(*
SPDX-FileCopyrightText: © 2026 Oleksandr Tiutyk <trofimich@gmail.com>
SPDX-License-Identifier: MIT
License: https://opensource.org/license/mit
*)

(*!
<summary>Provides STRING constants and helpers for text manipulation and value formatting.</summary>
<description>
Buffer ownership and size requirements are defined by each operation. ANY formatting reads the caller's value
through its type descriptor. Try methods contain exceptions; this does not validate buffer lifetime or undo
partial modifications.
Runtime type diagnostics use TYPE_ names for known classes and decimal codes for unknown values.
</description>
*)

{attribute 'no_explicit_call' := 'Direct call is not allowed'}
PROGRAM Strings
VAR_INPUT CONSTANT
	CharSize : BYTE := 1;
	//! <summary>ASCII space byte; values below it are control bytes in lexical text filters.</summary>
	ASCII_SPACE : BYTE := BYTE#16#20;
	NewLine : STRING(1) := '$R';
	Empty : STRING(0) := '';
	//! <summary>Standard three-dot ellipsis sequence for single-byte text truncation.</summary>
	ELLIPSIS : STRING(3) := '...';
END_VAR
VAR
	{attribute 'hide'} 
	_ClassName : STRING := __POUNAME();
END_VAR

(*!
<summary>Formats a supported ANY value as text of at most 255 characters.</summary>
<description>
Reads the borrowed live payload of supported types. Unsupported type classes produce a diagnostic marker
containing the type and size instead of interpreting the payload. The result is an independent bounded value.
</description>
*)
METHOD AnyToString : STRING(255)
VAR_INPUT
	value : ANY;
END_VAR
AnyToString := InternalAnyToString255(value := value);
END_METHOD

(*!
<summary>Formats a supported ANY value as text of at most 255 characters.</summary>
<description>
Reads the borrowed live payload of supported types. Unsupported type classes produce a diagnostic marker
containing the type and size instead of interpreting the payload. The result is an independent bounded value.
</description>
*)
METHOD AnyToString255 : STRING(255)
VAR_INPUT
	value : ANY;
END_VAR
AnyToString255 := InternalAnyToString255(value := value);
END_METHOD

(*!
<summary>
Formats a supported ANY value as text of at most 255 characters, fitting longer strings with an ellipsis
('...').
</summary>
<description>
Reads the borrowed live payload of supported types. String values longer than 255 characters are truncated to
252 characters and end with '...'. Non-string types and strings fitting in 255 characters are formatted
identically to AnyToString255.
</description>
<param name="value">Borrowed live value to format.</param>
*)
METHOD AnyToStringFit255 : STRING(255)
VAR_INPUT
	value : ANY;
END_VAR
VAR
	valueLength : UDINT;
END_VAR
AnyToStringFit255 := InternalAnyToString255(value := value);

IF value.TypeClass = __SYSTEM.TYPE_CLASS.TYPE_STRING THEN
	valueLength := InternalGetLength(value := value.pValue);

	IF valueLength > 255 THEN
		AnyToStringFit255 := Tc2_Standard.CONCAT(STR1 := Tc2_Standard.LEFT(STR := AnyToStringFit255, SIZE := 252), STR2 := '...');
	END_IF
ELSIF value.TypeClass = __SYSTEM.TYPE_CLASS.TYPE_WSTRING THEN
	valueLength := WideStrings.InternalGetLength(value := value.pValue);

	IF valueLength > 255 THEN
		AnyToStringFit255 := Tc2_Standard.CONCAT(STR1 := Tc2_Standard.LEFT(STR := AnyToStringFit255, SIZE := 252), STR2 := '...');
	END_IF
END_IF
END_METHOD

(*!
<summary>Appends one STRING to a caller-owned STRING buffer.</summary>
<description>
Requires live, null-terminated strings and a writable target whose declared size describes its capacity. After
validating the target type, an empty source completes without modifying the target. A non-STRING target raises
NotSupportedException; failure of the append helper raises TargetVariableMemoryOverflowException. Source
storage is borrowed only for this call.
Known runtime type classes appear by their TYPE_ names; unknown values retain their decimal codes.
</description>
*)
//!<param name="targetString">Writable STRING buffer to append to.</param>
//!<param name="sourceString">Text to append; empty leaves the target unchanged.</param>
METHOD Append
VAR_INPUT
	targetString : ANY_STRING;
END_VAR
VAR_IN_OUT CONSTANT
	sourceString : STRING;
END_VAR
VAR
	formattedExceptionMessage : WSTRING(255);
	
END_VAR
IF targetString.TypeClass <> __SYSTEM.TYPE_CLASS.TYPE_STRING THEN
	formattedExceptionMessage := Tc2_Utilities.WCONCAT(
		STR1 := "Not supported type ",
		STR2 := SystemTypeClassConvertor.ToWideString(typeClass := targetString.TypeClass)
	);

	Exceptions.ThrowNotSupported(
		sourceNamespaceName := NamespaceName,
		sourceClassName := ClassName,
		sourcePOUName := __POUNAME(),
		sourcePosition := __POSITION(),
		message := formattedExceptionMessage
	);
END_IF

IF sourceString = '' THEN
	RETURN;
END_IF

IF NOT InternalAppend(
	targetString := targetString,
	sourceString1 := ADR(sourceString),
	sourceString2 := 0,
	sourceString3 := 0,
	sourceString4 := 0,
	sourceString5 := 0,
	sourceString6 := 0,
	sourceString7 := 0,
	sourceString8 := 0,
	sourceString9 := 0,
	sourceString10 := 0
) THEN
	Exceptions.ThrowTargetVariableMemoryOverflow(
		sourceNamespaceName := NamespaceName,
		sourceClassName := ClassName,
		sourcePOUName := __POUNAME(),
		sourcePosition := __POSITION(),
		targetVariableName := 'targetString',
		targetVariableSize := TO_ULINT(targetString.diSize)
	); 
END_IF
END_METHOD

(*!
<summary>Appends up to ten STRING fragments in argument order, skipping empty fragments.</summary>
<description>
Requires live, null-terminated source strings and a writable STRING target with valid capacity metadata. Empty
fragments do not stop processing; if all are empty, the target is unchanged and the operation succeeds. Raises
NotSupportedException for a non-STRING target or TargetVariableMemoryOverflowException when appending fails.
Processing stops on the first append failure; earlier modifications are not rolled back. Source storage is
borrowed only for this call.
Known runtime type classes appear by their TYPE_ names; unknown values retain their decimal codes.
</description>
*)
METHOD Append255
VAR_INPUT
	targetString : ANY_STRING;
	sourceString1 : STRING(255);
	sourceString2 : STRING(255) := '';
	sourceString3 : STRING(255) := '';
	sourceString4 : STRING(255) := '';
	sourceString5 : STRING(255) := '';
	sourceString6 : STRING(255) := '';
	sourceString7 : STRING(255) := '';
	sourceString8 : STRING(255) := '';
	sourceString9 : STRING(255) := '';
	sourceString10 : STRING(255) := '';
END_VAR
VAR
	formattedExceptionMessage : WSTRING(255);
	
END_VAR
IF targetString.TypeClass <> __SYSTEM.TYPE_CLASS.TYPE_STRING THEN
	formattedExceptionMessage := Tc2_Utilities.WCONCAT(
		STR1 := "Not supported type ",
		STR2 := SystemTypeClassConvertor.ToWideString(typeClass := targetString.TypeClass)
	);

	Exceptions.ThrowNotSupported(
		sourceNamespaceName := NamespaceName,
		sourceClassName := ClassName,
		sourcePOUName := __POUNAME(),
		sourcePosition := __POSITION(),
		message := formattedExceptionMessage
	);
END_IF

	IF NOT InternalAppend(
		targetString := targetString,
		sourceString1 := ADR(sourceString1),
		sourceString2 := ADR(sourceString2),
		sourceString3 := ADR(sourceString3),
		sourceString4 := ADR(sourceString4),
		sourceString5 := ADR(sourceString5),
		sourceString6 := ADR(sourceString6),
		sourceString7 := ADR(sourceString7),
		sourceString8 := ADR(sourceString8),
		sourceString9 := ADR(sourceString9),
		sourceString10 := ADR(sourceString10)
	) THEN
	Exceptions.ThrowTargetVariableMemoryOverflow(
		sourceNamespaceName := NamespaceName,
		sourceClassName := ClassName,
		sourcePOUName := __POUNAME(),
		sourcePosition := __POSITION(),
		targetVariableName := 'targetString',
		targetVariableSize := TO_ULINT(targetString.diSize)
	); 
END_IF
END_METHOD

(*!
<summary>
Appends one STRING to a caller-owned STRING buffer, fitting available capacity with an ellipsis ('...') if
exceeded.
</summary>
<description>
Requires a writable STRING target with valid capacity metadata. If the appended text exceeds target capacity,
it is truncated so the final characters are '...' followed by a null-terminator. Raises NotSupportedException
for a non-STRING target. Source storage is borrowed only for this call.
Known runtime type classes appear by their TYPE_ names; unknown values retain their decimal codes.
</description>
<param name="targetString">Writable STRING buffer to append to.</param>
<param name="sourceString">Text to append; empty leaves the target unchanged.</param>
*)
METHOD AppendFit
VAR_INPUT
	targetString : ANY_STRING;
END_VAR
VAR_IN_OUT CONSTANT
	sourceString : STRING;
END_VAR
VAR
	formattedExceptionMessage : WSTRING(255);
END_VAR
IF targetString.TypeClass <> __SYSTEM.TYPE_CLASS.TYPE_STRING THEN
	formattedExceptionMessage := WideStrings.Concat255(
		"Not supported type ",
		SystemTypeClassConvertor.ToWideString(typeClass := targetString.TypeClass)
	);

	Exceptions.ThrowNotSupported(
		sourceNamespaceName := NamespaceName,
		sourceClassName := ClassName,
		sourcePOUName := __POUNAME(),
		sourcePosition := __POSITION(),
		message := formattedExceptionMessage
	);
END_IF

InternalAppendFit(targetString := targetString, sourceString := ADR(sourceString));
END_METHOD

(*!
<summary>
Appends up to ten STRING fragments in argument order, fitting available capacity with an ellipsis ('...') if
exceeded.
</summary>
<description>
Requires a writable STRING target with valid capacity metadata. Fragments are appended in order, skipping
empty fragments. If the combined text exceeds target capacity, it is truncated so the final characters are
'...' followed by a null-terminator. Raises NotSupportedException for a non-STRING target. Source storage is
borrowed only for this call.
Known runtime type classes appear by their TYPE_ names; unknown values retain their decimal codes.
</description>
<param name="targetString">Writable STRING buffer to append to.</param>
<param name="sourceString1">First text fragment to append.</param>
<param name="sourceString2">Second text fragment to append.</param>
<param name="sourceString3">Third text fragment to append.</param>
<param name="sourceString4">Fourth text fragment to append.</param>
<param name="sourceString5">Fifth text fragment to append.</param>
<param name="sourceString6">Sixth text fragment to append.</param>
<param name="sourceString7">Seventh text fragment to append.</param>
<param name="sourceString8">Eighth text fragment to append.</param>
<param name="sourceString9">Ninth text fragment to append.</param>
<param name="sourceString10">Tenth text fragment to append.</param>
*)
METHOD AppendFit255
VAR_INPUT
	targetString : ANY_STRING;
	sourceString1 : STRING(255);
	sourceString2 : STRING(255) := '';
	sourceString3 : STRING(255) := '';
	sourceString4 : STRING(255) := '';
	sourceString5 : STRING(255) := '';
	sourceString6 : STRING(255) := '';
	sourceString7 : STRING(255) := '';
	sourceString8 : STRING(255) := '';
	sourceString9 : STRING(255) := '';
	sourceString10 : STRING(255) := '';
END_VAR
VAR
	formattedExceptionMessage : WSTRING(255);
END_VAR
IF targetString.TypeClass <> __SYSTEM.TYPE_CLASS.TYPE_STRING THEN
	formattedExceptionMessage := Tc2_Utilities.WCONCAT(
		STR1 := "Not supported type ",
		STR2 := SystemTypeClassConvertor.ToWideString(typeClass := targetString.TypeClass)
	);

	Exceptions.ThrowNotSupported(
		sourceNamespaceName := NamespaceName,
		sourceClassName := ClassName,
		sourcePOUName := __POUNAME(),
		sourcePosition := __POSITION(),
		message := formattedExceptionMessage
	);
END_IF

InternalAppendFit(targetString := targetString, sourceString := ADR(sourceString1));

IF sourceString2 <> '' THEN
	InternalAppendFit(targetString := targetString, sourceString := ADR(sourceString2));
END_IF

IF sourceString3 <> '' THEN
	InternalAppendFit(targetString := targetString, sourceString := ADR(sourceString3));
END_IF

IF sourceString4 <> '' THEN
	InternalAppendFit(targetString := targetString, sourceString := ADR(sourceString4));
END_IF

IF sourceString5 <> '' THEN
	InternalAppendFit(targetString := targetString, sourceString := ADR(sourceString5));
END_IF

IF sourceString6 <> '' THEN
	InternalAppendFit(targetString := targetString, sourceString := ADR(sourceString6));
END_IF

IF sourceString7 <> '' THEN
	InternalAppendFit(targetString := targetString, sourceString := ADR(sourceString7));
END_IF

IF sourceString8 <> '' THEN
	InternalAppendFit(targetString := targetString, sourceString := ADR(sourceString8));
END_IF

IF sourceString9 <> '' THEN
	InternalAppendFit(targetString := targetString, sourceString := ADR(sourceString9));
END_IF

IF sourceString10 <> '' THEN
	InternalAppendFit(targetString := targetString, sourceString := ADR(sourceString10));
END_IF
END_METHOD

{attribute 'monitoring' := 'call'}
PROPERTY ClassName : REFERENCE TO STRING
GET
ClassName REF= _ClassName;
END_GET
END_PROPERTY

(*!
<summary>Concatenates up to sixteen text fragments without nested calls.</summary>
<description>
Fragments are appended in argument order. Empty and omitted optional fragments are skipped; they do not
prevent later fragments from being appended. The result is limited to 255 characters; excess text is truncated
by the standard concatenation function. No dynamic memory is allocated.
</description>
*)
METHOD Concat255 : STRING(255)
VAR_INPUT
	string1 : STRING(255);
	string2 : STRING(255);
	string3 : STRING(255) := '';
	string4 : STRING(255) := '';
	string5 : STRING(255) := '';
	string6 : STRING(255) := '';
	string7 : STRING(255) := '';
	string8 : STRING(255) := '';
	string9 : STRING(255) := '';
	string10 : STRING(255) := '';
	string11 : STRING(255) := '';
	string12 : STRING(255) := '';
	string13 : STRING(255) := '';
	string14 : STRING(255) := '';
	string15 : STRING(255) := '';
	string16 : STRING(255) := '';
END_VAR
Concat255 := Tc2_Standard.CONCAT(STR1 := string1, STR2 := string2);

IF Tc2_Standard.LEN(STR := string3) > 0 THEN
	Concat255 := Tc2_Standard.CONCAT(STR1 := Concat255, STR2 := string3);
END_IF

IF Tc2_Standard.LEN(STR := string4) > 0 THEN
	Concat255 := Tc2_Standard.CONCAT(STR1 := Concat255, STR2 := string4);
END_IF

IF Tc2_Standard.LEN(STR := string5) > 0 THEN
	Concat255 := Tc2_Standard.CONCAT(STR1 := Concat255, STR2 := string5);
END_IF

IF Tc2_Standard.LEN(STR := string6) > 0 THEN
	Concat255 := Tc2_Standard.CONCAT(STR1 := Concat255, STR2 := string6);
END_IF

IF Tc2_Standard.LEN(STR := string7) > 0 THEN
	Concat255 := Tc2_Standard.CONCAT(STR1 := Concat255, STR2 := string7);
END_IF

IF Tc2_Standard.LEN(STR := string8) > 0 THEN
	Concat255 := Tc2_Standard.CONCAT(STR1 := Concat255, STR2 := string8);
END_IF

IF Tc2_Standard.LEN(STR := string9) > 0 THEN
	Concat255 := Tc2_Standard.CONCAT(STR1 := Concat255, STR2 := string9);
END_IF

IF Tc2_Standard.LEN(STR := string10) > 0 THEN
	Concat255 := Tc2_Standard.CONCAT(STR1 := Concat255, STR2 := string10);
END_IF

IF Tc2_Standard.LEN(STR := string11) > 0 THEN
	Concat255 := Tc2_Standard.CONCAT(STR1 := Concat255, STR2 := string11);
END_IF

IF Tc2_Standard.LEN(STR := string12) > 0 THEN
	Concat255 := Tc2_Standard.CONCAT(STR1 := Concat255, STR2 := string12);
END_IF

IF Tc2_Standard.LEN(STR := string13) > 0 THEN
	Concat255 := Tc2_Standard.CONCAT(STR1 := Concat255, STR2 := string13);
END_IF

IF Tc2_Standard.LEN(STR := string14) > 0 THEN
	Concat255 := Tc2_Standard.CONCAT(STR1 := Concat255, STR2 := string14);
END_IF

IF Tc2_Standard.LEN(STR := string15) > 0 THEN
	Concat255 := Tc2_Standard.CONCAT(STR1 := Concat255, STR2 := string15);
END_IF

IF Tc2_Standard.LEN(STR := string16) > 0 THEN
	Concat255 := Tc2_Standard.CONCAT(STR1 := Concat255, STR2 := string16);
END_IF
END_METHOD

(*!
<summary>
Concatenates up to sixteen text fragments, fitting within 255 characters with an ellipsis ('...') if total
length is exceeded.
</summary>
<description>
Fragments are appended in argument order. Empty fragments are skipped. If the combined text exceeds 255
characters, the result is truncated to 252 characters and marked with a final '...'. No dynamic memory is
allocated.
</description>
<param name="string1">First text fragment.</param>
<param name="string2">Second text fragment.</param>
<param name="string3">Third text fragment.</param>
<param name="string4">Fourth text fragment.</param>
<param name="string5">Fifth text fragment.</param>
<param name="string6">Sixth text fragment.</param>
<param name="string7">Seventh text fragment.</param>
<param name="string8">Eighth text fragment.</param>
<param name="string9">Ninth text fragment.</param>
<param name="string10">Tenth text fragment.</param>
<param name="string11">Eleventh text fragment.</param>
<param name="string12">Twelfth text fragment.</param>
<param name="string13">Thirteenth text fragment.</param>
<param name="string14">Fourteenth text fragment.</param>
<param name="string15">Fifteenth text fragment.</param>
<param name="string16">Sixteenth text fragment.</param>
*)
METHOD ConcatFit255 : STRING(255)
VAR_INPUT
	string1 : STRING(255);
	string2 : STRING(255) := '';
	string3 : STRING(255) := '';
	string4 : STRING(255) := '';
	string5 : STRING(255) := '';
	string6 : STRING(255) := '';
	string7 : STRING(255) := '';
	string8 : STRING(255) := '';
	string9 : STRING(255) := '';
	string10 : STRING(255) := '';
	string11 : STRING(255) := '';
	string12 : STRING(255) := '';
	string13 : STRING(255) := '';
	string14 : STRING(255) := '';
	string15 : STRING(255) := '';
	string16 : STRING(255) := '';
END_VAR
VAR
	result : STRING(255);
	targetAny : __SYSTEM.AnyType;
END_VAR
targetAny.TypeClass := __SYSTEM.TYPE_CLASS.TYPE_STRING;
targetAny.pValue := ADR(result);
targetAny.diSize := SIZEOF(result);

InternalAppendFit(targetString := targetAny, sourceString := ADR(string1));

IF string2 <> '' THEN
	InternalAppendFit(targetString := targetAny, sourceString := ADR(string2));
END_IF

IF string3 <> '' THEN
	InternalAppendFit(targetString := targetAny, sourceString := ADR(string3));
END_IF

IF string4 <> '' THEN
	InternalAppendFit(targetString := targetAny, sourceString := ADR(string4));
END_IF

IF string5 <> '' THEN
	InternalAppendFit(targetString := targetAny, sourceString := ADR(string5));
END_IF

IF string6 <> '' THEN
	InternalAppendFit(targetString := targetAny, sourceString := ADR(string6));
END_IF

IF string7 <> '' THEN
	InternalAppendFit(targetString := targetAny, sourceString := ADR(string7));
END_IF

IF string8 <> '' THEN
	InternalAppendFit(targetString := targetAny, sourceString := ADR(string8));
END_IF

IF string9 <> '' THEN
	InternalAppendFit(targetString := targetAny, sourceString := ADR(string9));
END_IF

IF string10 <> '' THEN
	InternalAppendFit(targetString := targetAny, sourceString := ADR(string10));
END_IF

IF string11 <> '' THEN
	InternalAppendFit(targetString := targetAny, sourceString := ADR(string11));
END_IF

IF string12 <> '' THEN
	InternalAppendFit(targetString := targetAny, sourceString := ADR(string12));
END_IF

IF string13 <> '' THEN
	InternalAppendFit(targetString := targetAny, sourceString := ADR(string13));
END_IF

IF string14 <> '' THEN
	InternalAppendFit(targetString := targetAny, sourceString := ADR(string14));
END_IF

IF string15 <> '' THEN
	InternalAppendFit(targetString := targetAny, sourceString := ADR(string15));
END_IF

IF string16 <> '' THEN
	InternalAppendFit(targetString := targetAny, sourceString := ADR(string16));
END_IF

ConcatFit255 := result;
END_METHOD

(*!
<summary>Determines whether a string contains an exact, case-sensitive occurrence of a substring.</summary>
<description>
Returns TRUE when the substring is found. An empty search substring matches any source, including an empty
source. Returns FALSE when absent. Inputs must be live, null-terminated strings; they are borrowed only for
this call and are not modified.
</description>
<param name="stringToSearchIn">Text to search.</param>
<param name="stringToFind">Substring to locate; empty matches any string.</param>
*)
METHOD Contains : BOOL
VAR_IN_OUT CONSTANT
	stringToSearchIn : STRING;
	stringToFind : STRING;
END_VAR
Contains := Find(
	stringToSearchIn := stringToSearchIn,
	stringToFind := stringToFind
);
END_METHOD

(*!
<summary>Creates an enumerator over fragments of a borrowed source string.</summary>
<description>
The source must remain alive and unchanged during iteration. The splitter owns its current fragment; borrowed
fragment references expire on MoveNext, Reset or destruction. This method does not allocate the splitter with
__NEW. The initialized result has no fragment allocation until MoveNext; assigning it must not overwrite an
instance with an unreleased fragment. The caller is responsible for the result lifetime and cleanup, including
Reset when abandoning iteration. Do not copy an active splitter by value; use references. Only an instance
explicitly allocated with __NEW may be deleted with __DELETE.
</description>
*)
//!<param name="maxCount">
//! Maximum number of returned fragments; zero means unlimited. Empty fragments removed after optional
//! trimming do not count toward the limit. Remaining text is not returned after the limit is reached and is
//! not merged into the last fragment.
//! </param>
//!<param name="separator">
//! Copied separator containing 1 to 80 characters. An empty or longer value raises
//! ArgumentOutOfRangeException before initialization. The 255-character input capacity preserves rejection
//! of all values longer than 80.
//! </param>
METHOD CreateSplitter : StringSplittingEnumerator
VAR_IN_OUT CONSTANT
	sourceString : STRING;
END_VAR
VAR_INPUT
	separator : STRING(255);
	maxCount : UDINT := 0;
	trimEntries : BOOL := FALSE;
	removeEmptyEntries : BOOL := FALSE;
END_VAR
VAR
END_VAR
IF NOT __ISVALIDREF(sourceString) THEN
	Exceptions.ThrowArgumentNotSpecified(
		sourceNamespaceName := NamespaceName,
		sourceClassName := ClassName,
		sourcePOUName := __POUNAME(),
		sourcePosition := __POSITION(),
		argumentName := 'sourceString'
	);
END_IF

IF separator = '' OR_ELSE InternalGetLength(value := ADR(separator)) > 80 THEN
	Exceptions.ThrowArgumentOutOfRange(
		sourceNamespaceName := NamespaceName,
		sourceClassName := ClassName,
		sourcePOUName := __POUNAME(),
		sourcePosition := __POSITION(),
		argumentName := 'separator',
		argumentValue := separator
	);
END_IF

CreateSplitter.Initialize(
	sourceString := ADR(sourceString),
	separator := separator,
	maxCount := maxCount,
	trimEntries := trimEntries,
	removeEmptyEntries := removeEmptyEntries
);
END_METHOD

(*!
<summary>Finds the first exact, case-sensitive occurrence of a substring.</summary>
<description>
Returns TRUE with a one-based position when found. An empty search substring matches at position 1, including
in an empty source. Returns FALSE with position 0 when absent. Inputs must be live, null-terminated strings;
they are borrowed only for this call and are not modified.
</description>
*)
//!<param name="stringToSearchIn">Text to search.</param>
//!<param name="stringToFind">Substring to locate; empty matches at the beginning.</param>
//!<param name="position">One-based position in code units, or zero when absent.</param>
METHOD Find : BOOL
VAR_IN_OUT CONSTANT
	stringToSearchIn : STRING;
	stringToFind : STRING;
END_VAR
VAR_OUTPUT
	position : UDINT;
END_VAR
VAR
	stringToFindLength : UDINT;
END_VAR
position := 0;
stringToFindLength := InternalGetLength(value := ADR(stringToFind));

IF stringToFindLength = 0 THEN
	position := 1;
	Find := TRUE;
	RETURN;
END_IF

Find := InternalFind(
	stringToSearchIn := ADR(stringToSearchIn),
	stringToSearchInLength := InternalGetLength(value := ADR(stringToSearchIn)),
	stringToFind := ADR(stringToFind),
	stringToFindLength := stringToFindLength,
	position => position
);
END_METHOD

(*!
<summary>Returns the occupied byte size of terminated text.</summary>
<description>
Includes the terminating zero. This is the current text size, not the declared or allocated capacity; the
supplied string must remain valid during the call.
</description>
*)
METHOD GetActualSize : UDINT
VAR_IN_OUT CONSTANT
	value : STRING;
END_VAR
GetActualSize := InternalGetLength(value := ADR(value)) + CharSize;
END_METHOD

(*!
<summary>Returns the number of characters before the terminating zero.</summary>
<description>
Requires valid terminated text and excludes the terminator. Does not copy or modify the input.
</description>
*)
METHOD GetLength : UDINT
VAR_IN_OUT CONSTANT
	value : STRING;
END_VAR
GetLength := InternalGetLength(value := ADR(value));
END_METHOD

(*!
<summary>Formats a supported ANY value into a STRING of at most 255 characters.</summary>
<description>
Borrows the value storage for this call. The descriptor must identify a live value of the stated type. The
result does not retain a reference to the source. Unhandled type classes return a diagnostic marker containing
the type class and descriptor size in bytes, without reading value storage, allocating heap memory or raising
a formatting exception. This also applies to an unhandled type with a null data address.
Known runtime type classes appear by their TYPE_ names; unknown values retain their decimal codes.
</description>
<param name="value">Type descriptor and address of the value to format.</param>
*)
METHOD INTERNAL InternalAnyToString255 : STRING(255)
VAR_IN_OUT CONSTANT
	value : __SYSTEM.AnyType;
END_VAR
VAR
	anyBool : POINTER TO BOOL;

	anyByte : POINTER TO BYTE;
	anyWord : POINTER TO WORD;
	anyDWord : POINTER TO DWORD;
	anyLWord : POINTER TO LWORD;
	
	anySInt : POINTER TO SINT;
	anyInt : POINTER TO INT;
	anyDInt : POINTER TO DINT;
	anyLInt : POINTER TO LINT;
	
	anyUSInt : POINTER TO USINT;
	anyUInt : POINTER TO UINT;
	anyUDInt : POINTER TO UDINT;
	anyULInt : POINTER TO ULINT;
	
	anyReal : POINTER TO REAL;
	anyLReal : POINTER TO LREAL;

	anyString : POINTER TO STRING(255);
	anyWString : POINTER TO WSTRING(255);
	
	anyTime : POINTER TO TIME;
	anyLTime : POINTER TO LTIME;
	anyDate : POINTER TO DATE;
	anyDateAndTime : POINTER TO DATE_AND_TIME;
	anyTimeOfDay : POINTER TO TOD;

	anyPVoid : POINTER TO PVOID;
END_VAR
CASE value.TypeClass OF
	__SYSTEM.TYPE_CLASS.TYPE_BOOL:
		anyBool := value.pValue;
		InternalAnyToString255 := TO_STRING(anyBool^);		
	
	__SYSTEM.TYPE_CLASS.TYPE_BIT:
		anyByte := value.pValue;

		IF anyByte^ > 0 THEN
			InternalAnyToString255 := '1';		
		ELSE
			InternalAnyToString255 := '0';		
		END_IF
	
	__SYSTEM.TYPE_CLASS.TYPE_BYTE:
		anyByte := value.pValue;
		InternalAnyToString255 := TO_STRING(anyByte^);		
	__SYSTEM.TYPE_CLASS.TYPE_WORD:
		anyWord := value.pValue;
		InternalAnyToString255 := TO_STRING(anyWord^);
	__SYSTEM.TYPE_CLASS.TYPE_DWORD:
		anyDWord := value.pValue;
		InternalAnyToString255 := TO_STRING(anyDWord^);
	__SYSTEM.TYPE_CLASS.TYPE_LWORD:
		anyLWord := value.pValue;
		InternalAnyToString255 := TO_STRING(anyLWord^);
		
	__SYSTEM.TYPE_CLASS.TYPE_SINT:
		anySInt := value.pValue;
		InternalAnyToString255 := TO_STRING(anySInt^);
	__SYSTEM.TYPE_CLASS.TYPE_INT:
		anyInt := value.pValue;
		InternalAnyToString255 := TO_STRING(anyInt^);		
	__SYSTEM.TYPE_CLASS.TYPE_DINT:
		anyDInt := value.pValue;
		InternalAnyToString255 := TO_STRING(anyDInt^);
	__SYSTEM.TYPE_CLASS.TYPE_LINT:
		anyLInt := value.pValue;
		InternalAnyToString255 := TO_STRING(anyLInt^);
		
	__SYSTEM.TYPE_CLASS.TYPE_USINT:
		anyUSInt := value.pValue;
		InternalAnyToString255 := TO_STRING(anyUSInt^);
	__SYSTEM.TYPE_CLASS.TYPE_UINT:
		anyUInt := value.pValue;
		InternalAnyToString255 := TO_STRING(anyUInt^);		
	__SYSTEM.TYPE_CLASS.TYPE_UDINT:
		anyUDInt := value.pValue;
		InternalAnyToString255 := TO_STRING(anyUDInt^);
	__SYSTEM.TYPE_CLASS.TYPE_ULINT:
		anyULInt := value.pValue;
		InternalAnyToString255 := TO_STRING(anyULInt^);

	__SYSTEM.TYPE_CLASS.TYPE_REAL:
		anyReal := value.pValue;
		InternalAnyToString255 := TO_STRING(anyReal^);
	__SYSTEM.TYPE_CLASS.TYPE_LREAL:
		anyLReal := value.pValue;
		InternalAnyToString255 := TO_STRING(anyLReal^);
	
	__SYSTEM.TYPE_CLASS.TYPE_STRING:
		anyString := value.pValue;
		InternalAnyToString255 := anyString^;
	__SYSTEM.TYPE_CLASS.TYPE_WSTRING:
		anyWString := value.pValue;
		InternalAnyToString255 := TO_STRING(anyWString^);
	
	__SYSTEM.TYPE_CLASS.TYPE_TIME:
		anyTime := value.pValue;
		InternalAnyToString255 := TO_STRING(anyTime^);
	__SYSTEM.TYPE_CLASS.TYPE_LTIME:
		anyLTime := value.pValue;
		InternalAnyToString255 := TO_STRING(anyLTime^);
	__SYSTEM.TYPE_CLASS.TYPE_DATE:
		anyDate := value.pValue;
		InternalAnyToString255 := TO_STRING(anyDate^);
	__SYSTEM.TYPE_CLASS.TYPE_DATEANDTIME:
		anyDateAndTime := value.pValue;
		InternalAnyToString255 := TO_STRING(anyDateAndTime^);  
	__SYSTEM.TYPE_CLASS.TYPE_TIMEOFDAY:
		anyTimeOfDay := value.pValue;
		InternalAnyToString255 := TO_STRING(anyTimeOfDay^);
	
	__SYSTEM.TYPE_CLASS.TYPE_POINTER, __SYSTEM.TYPE_CLASS.TYPE_REFERENCE:
		anyPVoid := value.pValue;
		InternalAnyToString255 := Tc2_Utilities.PVOID_TO_HEXSTR(
			in := anyPVoid^,
			iPrecision := TO_INT(SIZEOF(PVOID) * 2),
			bLoCase := FALSE
		);		
	
	ELSE
		InternalAnyToString255 := Concat255(
			'<value unavailable; type class: ',
			SystemTypeClassConvertor.ToString(typeClass := value.TypeClass),
			'; size: ',
			TO_STRING(value.diSize),
			' bytes>'
		);
END_CASE
END_METHOD

(*!
<summary>Appends up to ten STRING fragments in argument order, skipping empty fragments.</summary>
<description>
Requires live, null-terminated source strings and a writable STRING target with valid capacity metadata. Empty
fragments do not stop processing; if all are empty, the target is unchanged and the operation succeeds.
Returns FALSE for a non-STRING target or when appending fails. Processing stops on the first append failure;
earlier modifications are not rolled back. Source storage is borrowed only for this call. Null source pointers
denote omitted fragments and are skipped.
</description>
*)
METHOD INTERNAL InternalAppend : BOOL
VAR_INPUT
	targetString : __SYSTEM.AnyType;
	sourceString1 : POINTER TO STRING;
	sourceString2 : POINTER TO STRING;
	sourceString3 : POINTER TO STRING;
	sourceString4 : POINTER TO STRING;
	sourceString5 : POINTER TO STRING;
	sourceString6 : POINTER TO STRING;
	sourceString7 : POINTER TO STRING;
	sourceString8 : POINTER TO STRING;
	sourceString9 : POINTER TO STRING;
	sourceString10 : POINTER TO STRING;
END_VAR
InternalAppend := FALSE;

IF targetString.TypeClass <> __SYSTEM.TYPE_CLASS.TYPE_STRING THEN
	RETURN;
END_IF

IF sourceString1 <> 0 AND_THEN Tc2_Utilities.LEN2(pSTRING := sourceString1) > 0 THEN
	IF NOT Tc2_Utilities.CONCAT2(
		pSrcString1 := targetString.pValue,
		pSrcString2 := sourceString1,
		pDstString := targetString.pValue,
		nDstSize := TO_UDINT(targetString.diSize)
	) THEN
		RETURN;
	END_IF
END_IF

IF sourceString2 <> 0 AND_THEN Tc2_Utilities.LEN2(pSTRING := sourceString2) > 0 THEN
	IF NOT Tc2_Utilities.CONCAT2(
		pSrcString1 := targetString.pValue,
		pSrcString2 := sourceString2,
		pDstString := targetString.pValue,
		nDstSize := TO_UDINT(targetString.diSize)
	) THEN
		RETURN;
	END_IF
END_IF

IF sourceString3 <> 0 AND_THEN Tc2_Utilities.LEN2(pSTRING := sourceString3) > 0 THEN
	IF NOT Tc2_Utilities.CONCAT2(
		pSrcString1 := targetString.pValue,
		pSrcString2 := sourceString3,
		pDstString := targetString.pValue,
		nDstSize := TO_UDINT(targetString.diSize)
	) THEN
		RETURN;
	END_IF
END_IF

IF sourceString4 <> 0 AND_THEN Tc2_Utilities.LEN2(pSTRING := sourceString4) > 0 THEN
	IF NOT Tc2_Utilities.CONCAT2(
		pSrcString1 := targetString.pValue,
		pSrcString2 := sourceString4,
		pDstString := targetString.pValue,
		nDstSize := TO_UDINT(targetString.diSize)
	) THEN
		RETURN;
	END_IF
END_IF

IF sourceString5 <> 0 AND_THEN Tc2_Utilities.LEN2(pSTRING := sourceString5) > 0 THEN
	IF NOT Tc2_Utilities.CONCAT2(
		pSrcString1 := targetString.pValue,
		pSrcString2 := sourceString5,
		pDstString := targetString.pValue,
		nDstSize := TO_UDINT(targetString.diSize)
	) THEN
		RETURN;
	END_IF
END_IF

IF sourceString6 <> 0 AND_THEN Tc2_Utilities.LEN2(pSTRING := sourceString6) > 0 THEN
	IF NOT Tc2_Utilities.CONCAT2(
		pSrcString1 := targetString.pValue,
		pSrcString2 := sourceString6,
		pDstString := targetString.pValue,
		nDstSize := TO_UDINT(targetString.diSize)
	) THEN
		RETURN;
	END_IF
END_IF

IF sourceString7 <> 0 AND_THEN Tc2_Utilities.LEN2(pSTRING := sourceString7) > 0 THEN
	IF NOT Tc2_Utilities.CONCAT2(
		pSrcString1 := targetString.pValue,
		pSrcString2 := sourceString7,
		pDstString := targetString.pValue,
		nDstSize := TO_UDINT(targetString.diSize)
	) THEN
		RETURN;
	END_IF
END_IF

IF sourceString8 <> 0 AND_THEN Tc2_Utilities.LEN2(pSTRING := sourceString8) > 0 THEN
	IF NOT Tc2_Utilities.CONCAT2(
		pSrcString1 := targetString.pValue,
		pSrcString2 := sourceString8,
		pDstString := targetString.pValue,
		nDstSize := TO_UDINT(targetString.diSize)
	) THEN
		RETURN;
	END_IF
END_IF

IF sourceString9 <> 0 AND_THEN Tc2_Utilities.LEN2(pSTRING := sourceString9) > 0 THEN
	IF NOT Tc2_Utilities.CONCAT2(
		pSrcString1 := targetString.pValue,
		pSrcString2 := sourceString9,
		pDstString := targetString.pValue,
		nDstSize := TO_UDINT(targetString.diSize)
	) THEN
		RETURN;
	END_IF
END_IF

IF sourceString10 <> 0 AND_THEN Tc2_Utilities.LEN2(pSTRING := sourceString10) > 0 THEN
	IF NOT Tc2_Utilities.CONCAT2(
		pSrcString1 := targetString.pValue,
		pSrcString2 := sourceString10,
		pDstString := targetString.pValue,
		nDstSize := TO_UDINT(targetString.diSize)
	) THEN
		RETURN;
	END_IF
END_IF

InternalAppend := TRUE;
END_METHOD

(*!
<summary>Appends text to a STRING buffer, marking truncation when capacity permits.</summary>
<description>
Requires live, terminated input and writable target storage of the matching encoding.
On overflow, capacities of at least three characters use three dots. Capacities of one or two use one dot.
A buffer with room only for its terminator stays empty and succeeds. Missing terminator space or an invalid
target returns FALSE. The caller handles native exceptions.
</description>
*)
METHOD INTERNAL InternalAppendFit : BOOL
VAR_INPUT
	targetString : __SYSTEM.AnyType;
	sourceString : POINTER TO STRING;
END_VAR
VAR
	maxCapacity : UDINT;
	currentLength : UDINT;
	sourceLength : UDINT;
	availableChars : UDINT;
	targetBytes : POINTER TO BYTE;
END_VAR
InternalAppendFit := FALSE;

IF targetString.TypeClass <> __SYSTEM.TYPE_CLASS.TYPE_STRING
	OR_ELSE targetString.pValue = 0
	OR_ELSE targetString.diSize < 1
THEN
	RETURN;
END_IF

IF sourceString = 0 THEN
	InternalAppendFit := TRUE;
	RETURN;
END_IF

sourceLength := TO_UDINT(Tc2_Utilities.LEN2(pSTRING := sourceString));

IF sourceLength = 0 THEN
	InternalAppendFit := TRUE;
	RETURN;
END_IF

maxCapacity := TO_UDINT(targetString.diSize) - 1;
currentLength := TO_UDINT(Tc2_Utilities.LEN2(pSTRING := targetString.pValue));

IF currentLength > maxCapacity THEN
	currentLength := maxCapacity;
END_IF

targetBytes := targetString.pValue;

IF currentLength + sourceLength <= maxCapacity THEN
	InternalAppendFit := Tc2_Utilities.CONCAT2(
		pSrcString1 := targetString.pValue,
		pSrcString2 := sourceString,
		pDstString := targetString.pValue,
		nDstSize := TO_UDINT(targetString.diSize)
	);

	RETURN;
ELSE
	IF maxCapacity >= 3 THEN
		IF currentLength >= maxCapacity - 3 THEN
			currentLength := maxCapacity - 3;
			availableChars := 0;
		ELSE
			availableChars := maxCapacity - 3 - currentLength;
			Tc2_System.MEMCPY(destAddr := targetString.pValue + currentLength, srcAddr := sourceString, n := availableChars);
		END_IF

		targetBytes[currentLength + availableChars] := 16#2E; // '.'
		targetBytes[currentLength + availableChars + 1] := 16#2E; // '.'
		targetBytes[currentLength + availableChars + 2] := 16#2E; // '.'
		targetBytes[currentLength + availableChars + 3] := 0;
	ELSIF maxCapacity > 0 THEN
		IF currentLength >= maxCapacity - 1 THEN
			currentLength := maxCapacity - 1;
		END_IF
		
		targetBytes[currentLength] := 16#2E;
		targetBytes[currentLength + 1] := 0;
	ELSE
		targetBytes[0] := 0;
	END_IF
END_IF

InternalAppendFit := TRUE;
END_METHOD

(*!
<summary>Finds the first exact occurrence of a nonempty substring in buffers with supplied lengths.</summary>
<description>
Lengths and the one-based result position are measured in code units, excluding terminators. Caller-provided
lengths must describe accessible buffers. Returns FALSE and position 0 for an empty search substring or no
match. Unlike public Find, this helper does not match an empty substring, allowing replacement and splitting
loops to make progress.
</description>
*)
METHOD INTERNAL InternalFind : BOOL
VAR_INPUT
	stringToSearchIn : POINTER TO STRING;
	stringToSearchInLength : UDINT;
	stringToFind : POINTER TO STRING;
	stringToFindLength : UDINT;
END_VAR
VAR_OUTPUT
	position : UDINT;
END_VAR
VAR	
	i : UDINT;
END_VAR
InternalFind := FALSE;
position := 0;

IF stringToFindLength = 0 OR_ELSE stringToSearchInLength < stringToFindLength THEN
	RETURN;
END_IF

FOR i := 0 TO stringToSearchInLength - stringToFindLength DO
	IF Tc2_System.MEMCMP(pBuf1 := stringToSearchIn + i, pBuf2 := stringToFind, n := stringToFindLength * CharSize) = 0 THEN
		position := i + 1;
		InternalFind := TRUE;
		RETURN;
	END_IF
END_FOR
END_METHOD

(*!
<summary>Returns the length of text at the supplied address.</summary>
<description>
Returns zero for a null address. A nonzero address must point to readable, correctly terminated text; this
method does not establish pointer validity or buffer capacity.
</description>
*)
METHOD INTERNAL InternalGetLength : UDINT
VAR_INPUT
	value : POINTER TO STRING;
END_VAR
InternalGetLength := SEL(value = 0, Tc2_Utilities.LEN2(pSTRING := value), 0);
END_METHOD

(*!
<summary>Builds joined text from the selected enumerated values in the supplied buffer.</summary>
<description>
Clears the target before joining and consumes the enumerator from its current position. Strings of the target
encoding use a borrowed reference regardless of their byte size. Other types use AsString255 and a matching
255-character local buffer, with that conversion method's truncation and exception behavior. Returns FALSE on
an incompatible target or append failure; partial text is not rolled back. Referenced data must remain valid
during each append. A latched allocation failure stops enumeration and returns FALSE.
</description>
*)
METHOD INTERNAL InternalJoin : BOOL
VAR_INPUT
	targetString : __SYSTEM.AnyType;
	separator : POINTER TO STRING;
	sourceEnumerator : IEnumerator;
	startIndex : UDINT;
	count : UDINT;
END_VAR
VAR
	currentValue : REFERENCE TO GENERIC_VALUE;
	string255 : STRING(255);
	stringReference : REFERENCE TO STRING;
	currentCount : UDINT;
	currentIndex : UDINT;
END_VAR
IF DynamicMemoryManager.HasAllocationFailed THEN
	RETURN;
END_IF

IF targetString.TypeClass <> __SYSTEM.TYPE_CLASS.TYPE_STRING THEN
	RETURN;
END_IF

Tc2_System.MEMSET(destAddr := targetString.pValue, fillByte := 0, n := TO_UDINT(targetString.diSize));

InternalJoin := TRUE;

WHILE NOT DynamicMemoryManager.HasAllocationFailed AND_THEN sourceEnumerator.MoveNext() DO
	IF DynamicMemoryManager.HasAllocationFailed THEN
		EXIT;
	END_IF

	currentValue REF= sourceEnumerator.Current;

	IF DynamicMemoryManager.HasAllocationFailed THEN
		EXIT;
	END_IF
	
	IF NOT __ISVALIDREF(currentValue) OR_ELSE currentIndex < startIndex THEN
		currentIndex := currentIndex + 1;
   		CONTINUE;
	END_IF
	
	IF currentCount > 0 THEN
		InternalJoin := InternalJoin AND Tc2_Utilities.CONCAT2(
			targetString.pValue,
			separator,
			targetString.pValue,
			TO_UDINT(targetString.diSize)
		);		
	END_IF

	IF NOT InternalJoin THEN
		RETURN;
	END_IF
		
	IF currentValue.TypeClass = GENERIC_TYPE_CLASS.STRING_8 THEN
		stringReference REF= currentValue.AsStringReference();

		InternalJoin := InternalJoin AND Tc2_Utilities.CONCAT2(
			targetString.pValue,
			ADR(stringReference),
			targetString.pValue,
			TO_UDINT(targetString.diSize)
		);
	ELSE
		string255 := currentValue.AsString255();

		InternalJoin := InternalJoin AND Tc2_Utilities.CONCAT2(
			targetString.pValue,
			ADR(string255),
			targetString.pValue,
			TO_UDINT(targetString.diSize)
		);
	END_IF
	
	IF NOT InternalJoin THEN
		RETURN;
	END_IF

	currentCount := currentCount + 1;
	currentIndex := currentIndex + 1;
	
	IF count > 0 AND_THEN currentCount >= count THEN
		EXIT;
	END_IF	
END_WHILE

InternalJoin := InternalJoin AND NOT DynamicMemoryManager.HasAllocationFailed;
END_METHOD

(*!
<summary>Replaces matching substrings in the supplied text buffer.</summary>
<description>
Replaces exact, case-sensitive, non-overlapping occurrences in place. An empty oldSubstring succeeds without
changes and sets replacementCount to zero. An empty newSubstring deletes matched text. Zero maxReplacements
means no replacement limit; skipReplacements skips the first matching occurrences. Returns FALSE if a memory
operation fails or the result does not fit. Replacement is not atomic. If the next replacement would exceed
buffer capacity, it is not performed; completed replacements remain, replacementCount reports their count, and
the valid source remains null-terminated. These guarantees concern capacity failure with valid input buffers,
not invalid memory access. The caller supplies live buffers of the correct encoding; sourceString must be
writable and its size must include space for the terminator.
</description>
*)
//!<param name="oldSubstring">Text to replace; empty performs no replacements.</param>
//!<param name="newSubstring">Replacement text; empty deletes each selected match.</param>
//!<param name="replacementCount">Number of completed replacements.</param>
METHOD INTERNAL InternalReplaceInSource : BOOL
VAR_INPUT
	sourceString : __SYSTEM.AnyType;
	oldSubstring : POINTER TO STRING;
	newSubstring : POINTER TO STRING;
	maxReplacements : UINT;
	skipReplacements : UINT;
END_VAR
VAR_OUTPUT
	replacementCount : UINT;
END_VAR
VAR
	sourceStringMemorySize : UDINT;
	sourceStringLength : UDINT;

	handledString : POINTER TO STRING;
	handledStringLength : UDINT;
		
	oldSubstringLength : UDINT;
	newSubstringLength : UDINT;
	checkMemorySize : BOOL;	
	
	substringPosition : UDINT;

	skipCount : UINT;
	
	memFunctionResult : UDINT;
END_VAR
InternalReplaceInSource := FALSE;
replacementCount := 0;
oldSubstringLength := InternalGetLength(value := oldSubstring);

IF oldSubstringLength = 0 THEN
	InternalReplaceInSource := TRUE;
	RETURN;
END_IF

sourceStringMemorySize := TO_UDINT(sourceString.diSize);
sourceStringLength := InternalGetLength(value := sourceString.pValue);

handledString := sourceString.pValue;
handledStringLength := sourceStringLength;

newSubstringLength := InternalGetLength(value := newSubstring);
checkMemorySize := oldSubstringLength < newSubstringLength;

WHILE handledStringLength >= oldSubstringLength DO
	IF NOT InternalFind(
		stringToSearchIn := handledString,
		stringToSearchInLength := handledStringLength / CharSize,
		stringToFind := oldSubstring,
		stringToFindLength := oldSubstringLength / CharSize,
		position => substringPosition
	) THEN
		EXIT;
	END_IF
	
	IF skipReplacements > 0 AND_THEN skipCount < skipReplacements THEN
		skipCount := skipCount + 1;

		handledString := handledString + oldSubstringLength + (substringPosition * CharSize) - CharSize;	
		handledStringLength := handledStringLength - oldSubstringLength - (substringPosition * CharSize) + CharSize;
		
		CONTINUE;		
	END_IF
	
	handledString := handledString + (substringPosition * CharSize) - CharSize;
	handledStringLength := handledStringLength - (substringPosition * CharSize) + CharSize;

	sourceStringLength := sourceStringLength + newSubstringLength - oldSubstringLength;
	
	IF checkMemorySize AND_THEN sourceStringLength + CharSize > sourceStringMemorySize THEN
		RETURN;
	END_IF
	
	IF oldSubstringLength <> newSubstringLength THEN
		memFunctionResult := Tc2_System.MEMMOVE(
			destAddr := handledString + newSubstringLength,
			srcAddr := handledString + oldSubstringLength,
			n := handledStringLength - oldSubstringLength + CharSize
		);
		
		IF memFunctionResult < 1 THEN
			RETURN;			
		END_IF
		
		handledStringLength := handledStringLength + newSubstringLength - oldSubstringLength;
	END_IF
	
	IF newSubstringLength > 0 THEN
		memFunctionResult := Tc2_System.MEMCPY(destAddr := handledString, srcAddr := newSubstring, n := newSubstringLength);
	
		IF memFunctionResult < 1 THEN
			RETURN;			
		END_IF		
	END_IF
	
	replacementCount := replacementCount + 1;
	
	IF maxReplacements > 0 AND_THEN replacementCount>= maxReplacements THEN
		EXIT;
	END_IF

	handledString := handledString + newSubstringLength;	
	handledStringLength := handledStringLength - newSubstringLength;
END_WHILE

InternalReplaceInSource := TRUE;
END_METHOD

(*!
<summary>Checks the complete input text for floating-point syntax.</summary>
<description>
Accepts decimal digits with an optional leading sign, at most one decimal point before an optional e/E
exponent, and an optional sign immediately after the exponent marker. Requires a mantissa digit and, when an
exponent is present, an exponent digit. Empty strings, whitespace and other characters are rejected. This is a
lexical check, not a numeric range or representability check. The caller supplies a live null-terminated
string, borrowed read-only for the call; processing is not limited to 255 characters and its cost grows with
input length.
</description>
*)
//!<param name="stringToCheck">Complete text to validate.</param>
METHOD IsFloat : BOOL
VAR_IN_OUT CONSTANT
    stringToCheck : STRING;
END_VAR
VAR
    i : UDINT;
    stringLength : UDINT;

    digitFound : BOOL;
    dotFound : BOOL;
    exponentFound : BOOL;
    exponentDigitFound : BOOL;
END_VAR
IsFloat := FALSE;
stringLength := Tc2_Utilities.LEN2(pSTRING := ADR(stringToCheck));

IF stringLength = 0 THEN
	RETURN;
END_IF

FOR i := 0 TO stringLength - 1 DO
    // sign can be first character 
    IF i = 0 AND_THEN (stringToCheck[i] = 43 OR_ELSE stringToCheck[i] = 45) THEN
        CONTINUE;
    END_IF

    // digit 
    IF stringToCheck[i] >= 48 AND_THEN stringToCheck[i] <= 57 THEN
        IF exponentFound THEN
            exponentDigitFound := TRUE;
        ELSE
            digitFound := TRUE;
        END_IF
		
        CONTINUE;
    END_IF

    // decimal point 
    IF stringToCheck[i] = 46 THEN
        IF dotFound OR exponentFound THEN
            RETURN;
        END_IF
		
        dotFound := TRUE;
		
        CONTINUE;
    END_IF

    // exponent
    IF stringToCheck[i] = 69 OR_ELSE stringToCheck[i] = 101 THEN
        IF exponentFound OR NOT digitFound THEN
            RETURN;
        END_IF
		
        exponentFound := TRUE;
		
        CONTINUE;
    END_IF

    // sign after e/E 
    IF exponentFound AND_THEN (stringToCheck[i] = 43 OR_ELSE stringToCheck[i] = 45) THEN
        IF stringToCheck[i - 1] = 69 OR_ELSE stringToCheck[i - 1] = 101 THEN
            CONTINUE;
        ELSE
            RETURN;
        END_IF
    END_IF

    // invalid symbol 
    RETURN;
END_FOR

IF exponentFound THEN
    IsFloat := digitFound AND_THEN exponentDigitFound;
ELSE
    IsFloat := digitFound;
END_IF
END_METHOD

(*!
<summary>Checks the complete input text for signed integer syntax.</summary>
<description>
Accepts decimal digits with an optional leading plus or minus sign; at least one digit is required. Empty
strings, whitespace and other characters are rejected. This is a lexical check, not a numeric range or
representability check. The caller supplies a live null-terminated string, borrowed read-only for the call;
processing is not limited to 255 characters and its cost grows with input length.
</description>
*)
//!<param name="stringToCheck">Complete text to validate.</param>
METHOD IsInteger : BOOL
VAR_IN_OUT CONSTANT
    stringToCheck : STRING;
END_VAR
VAR
    i : UDINT;
    stringLength : UDINT;

    digitFound : BOOL;
END_VAR
IsInteger := FALSE;
stringLength := Tc2_Utilities.LEN2(pSTRING := ADR(stringToCheck));

IF stringLength = 0 THEN
	RETURN;
END_IF

FOR i := 0 TO stringLength - 1 DO
    // sign can be first character 
    IF i = 0 AND_THEN (stringToCheck[i] = 43 OR_ELSE stringToCheck[i] = 45) THEN
        CONTINUE;
    END_IF

    // digit 
    IF stringToCheck[i] >= 48 AND_THEN stringToCheck[i] <= 57 THEN
		digitFound := TRUE;
		
        CONTINUE;
    END_IF

    // invalid symbol 
    RETURN;
END_FOR

IsInteger := digitFound;
END_METHOD

(*!
<summary>Reports whether the reference is absent, empty or contains only recognized whitespace.</summary>
<description>
A valid reference must designate readable terminated text. Uses the whitespace characters explicitly
recognized by this implementation; does not validate arbitrary addresses or normalize text.
</description>
*)
METHOD IsNullOrWhiteSpace : BOOL
VAR_INPUT
	stringToCheck : REFERENCE TO STRING;
END_VAR
VAR
	i : DINT;
	
	stringData : POINTER TO BYTE;
END_VAR
IsNullOrWhiteSpace := TRUE;

IF NOT __ISVALIDREF(stringToCheck) THEN
	RETURN;
END_IF

stringData := ADR(stringToCheck);

WHILE stringData[i] <> 0 DO
	CASE stringData[i] OF
		16#20, 16#09, 16#0A, 16#0B, 16#0C, 16#0D:
			i := i + 1;
			
		ELSE
			IsNullOrWhiteSpace := FALSE;
			RETURN;
	END_CASE 
END_WHILE
END_METHOD

(*!
<summary>Checks the complete input text for unsigned integer syntax.</summary>
<description>
Accepts decimal digits with an optional leading plus sign; at least one digit is required. Empty strings,
whitespace and other characters are rejected. This is a lexical check, not a numeric range or representability
check. The caller supplies a live null-terminated string, borrowed read-only for the call; processing is not
limited to 255 characters and its cost grows with input length.
</description>
*)
//!<param name="stringToCheck">Complete text to validate.</param>
METHOD IsUnsignedInteger : BOOL
VAR_IN_OUT CONSTANT
    stringToCheck : STRING;
END_VAR
VAR
    i : UDINT;
    stringLength : UDINT;

    digitFound : BOOL;
END_VAR
IsUnsignedInteger := FALSE;
stringLength := Tc2_Utilities.LEN2(pSTRING := ADR(stringToCheck));

IF stringLength = 0 THEN
	RETURN;
END_IF

FOR i := 0 TO stringLength - 1 DO
    // + can be first character 
    IF i = 0 AND_THEN stringToCheck[i] = 43 THEN
        CONTINUE;
    END_IF

    // digit 
    IF stringToCheck[i] >= 48 AND_THEN stringToCheck[i] <= 57 THEN
		digitFound := TRUE;
		
        CONTINUE;
    END_IF

    // invalid symbol 
    RETURN;
END_FOR

IsUnsignedInteger := digitFound;
END_METHOD

(*!
<summary>Joins selected enumerated values into the supplied STRING buffer with a separator.</summary>
<description>
Validates the target string type and a non-null enumerator, then clears the target and advances the enumerator
from its current position without resetting it. Invalid Current references are skipped. Inserts separators
between included values, including empty text values. Does not dispose or retain the enumerator; its lifetime
remains the caller's responsibility. Raises NotSupportedException for the wrong target type,
ArgumentNotSpecifiedException for a null enumerator and TargetVariableMemoryOverflowException on append
failure. A latched allocation failure is raised before reporting append failure.
Enumerator and conversion exceptions propagate. Partial text and the advanced enumerator position are
not rolled back. The caller supplies live writable target storage and source data that remain valid during the
operation. Strings of the target encoding are joined through a borrowed reference without a 255-character
intermediate limit. Other values use AsString255 with its default conversion policy and 255-character
capacity; unsupported conversions raise an exception.
Known runtime type classes appear by their TYPE_ names; unknown values retain their decimal codes.
</description>
*)
//!<param name="targetString">
//! Destination buffer, including capacity for the terminator; previous contents are cleared after argument
//! validation.
//! </param>
//!<param name="separator">Text inserted between included values.</param>
//!<param name="sourceEnumerator">Borrowed enumerator, consumed by MoveNext without Reset.</param>
//!<param name="startIndex">
//! Number of positions to skip among subsequent MoveNext results, including invalid Current references.
//! </param>
//!<param name="count">Maximum number of included values; zero consumes all remaining eligible values.</param>
METHOD Join
VAR_INPUT
	targetString : ANY_STRING;
END_VAR
VAR_INPUT
	separator : STRING;
	sourceEnumerator : IEnumerator;
	startIndex : UDINT := 0;
	count : UDINT := 0;
END_VAR
VAR
	formattedExceptionMessage : WSTRING(255);
	
END_VAR
IF targetString.TypeClass <> __SYSTEM.TYPE_CLASS.TYPE_STRING THEN
	formattedExceptionMessage := Tc2_Utilities.WCONCAT(
		STR1 := "Not supported type ",
		STR2 := SystemTypeClassConvertor.ToWideString(typeClass := targetString.TypeClass)
	);

	Exceptions.ThrowNotSupported(
		sourceNamespaceName := NamespaceName,
		sourceClassName := ClassName,
		sourcePOUName := __POUNAME(),
		sourcePosition := __POSITION(),
		message := formattedExceptionMessage
	);
END_IF

IF sourceEnumerator = 0 THEN
	Exceptions.ThrowArgumentNotSpecified(
		sourceNamespaceName := NamespaceName,
		sourceClassName := ClassName,
		sourcePOUName := __POUNAME(),
		sourcePosition := __POSITION(),
		argumentName := 'sourceEnumerator'
	);
END_IF

IF NOT InternalJoin(
	targetString := targetString,
	separator := ADR(separator),
	sourceEnumerator := sourceEnumerator,
	startIndex := startIndex,
	count := count
) THEN
	DynamicMemoryManager.RaiseIfAllocationFailed();

	Exceptions.ThrowTargetVariableMemoryOverflow(
		sourceNamespaceName := NamespaceName,
		sourceClassName := ClassName,
		sourcePOUName := __POUNAME(),
		sourcePosition := __POSITION(),
		targetVariableName := 'targetString',
		targetVariableSize := TO_ULINT(targetString.diSize)
	); 
END_IF
END_METHOD

(*!
<summary>Provides the library namespace used in diagnostics.</summary>
<description>
Borrowed read-only reference to the compiler-initialized library namespace; no ownership transfer.
</description>
*)
{attribute 'monitoring' := 'call'}
PROPERTY NamespaceName : REFERENCE TO STRING
GET
NamespaceName REF= CurrentNamespace.Name;
END_GET
END_PROPERTY

(*!
<summary>Replaces matching substrings in the supplied text buffer.</summary>
<description>
Replaces exact, case-sensitive, non-overlapping occurrences in place. An empty oldSubstring succeeds without
changes and sets replacementCount to zero. An empty newSubstring deletes matched text. Zero maxReplacements
means no replacement limit; skipReplacements skips the first matching occurrences. Raises
NotSupportedException for an incompatible source type and TargetVariableMemoryOverflowException if replacement
cannot complete. Replacement is not atomic. If the next replacement would exceed buffer capacity, it is not
performed; completed replacements remain, replacementCount reports their count, and the valid source remains
null-terminated. These guarantees concern capacity failure with valid input buffers, not invalid memory
access. The caller supplies live buffers of the correct encoding; sourceString must be writable and its size
must include space for the terminator.
Known runtime type classes appear by their TYPE_ names; unknown values retain their decimal codes.
</description>
*)
//!<param name="oldSubstring">Text to replace; empty performs no replacements.</param>
//!<param name="newSubstring">Replacement text; empty deletes each selected match.</param>
//!<param name="replacementCount">Number of completed replacements.</param>
METHOD ReplaceInSource
VAR_INPUT
	sourceString : ANY_STRING;
END_VAR
VAR_IN_OUT CONSTANT
	oldSubstring : STRING;
	newSubstring : STRING;
END_VAR
VAR_INPUT
	maxReplacements : UINT := 0;
	skipReplacements : UINT := 0;
END_VAR
VAR_OUTPUT
	replacementCount : UINT;
END_VAR
VAR	
	
	replaceResult : BOOL; 
END_VAR
VAR
	formattedExceptionMessage : WSTRING(255);
END_VAR
IF sourceString.TypeClass <> __SYSTEM.TYPE_CLASS.TYPE_STRING THEN
	formattedExceptionMessage := Tc2_Utilities.WCONCAT(
		STR1 := "Not supported type ",
		STR2 := SystemTypeClassConvertor.ToWideString(typeClass := sourceString.TypeClass)
	);

	Exceptions.ThrowNotSupported(
		sourceNamespaceName := NamespaceName,
		sourceClassName := ClassName,
		sourcePOUName := __POUNAME(),
		sourcePosition := __POSITION(),
		message := formattedExceptionMessage
	);
END_IF

IF NOT InternalReplaceInSource(
	sourceString := sourceString,
	oldSubstring := ADR(oldSubstring),
	newSubstring := ADR(newSubstring),
	maxReplacements := maxReplacements,
	skipReplacements := skipReplacements,
	replacementCount => replacementCount
) THEN
	Exceptions.ThrowTargetVariableMemoryOverflow(
		sourceNamespaceName := NamespaceName,
		sourceClassName := ClassName,
		sourcePOUName := __POUNAME(),
		sourcePosition := __POSITION(),
		targetVariableName := 'sourceString',
		targetVariableSize := TO_UDINT(sourceString.diSize)
	);
END_IF
END_METHOD

(*!
<summary>Replaces matching substrings in the supplied text buffer.</summary>
<description>
Replaces exact, case-sensitive, non-overlapping occurrences in place. An empty oldSubstring succeeds without
changes and sets replacementCount to zero. An empty newSubstring deletes matched text. Zero maxReplacements
means no replacement limit; skipReplacements skips the first matching occurrences. Raises
NotSupportedException for an incompatible source type and TargetVariableMemoryOverflowException if replacement
cannot complete. Replacement is not atomic. If the next replacement would exceed buffer capacity, it is not
performed; completed replacements remain, replacementCount reports their count, and the valid source remains
null-terminated. These guarantees concern capacity failure with valid input buffers, not invalid memory
access. The caller supplies live buffers of the correct encoding; sourceString must be writable and its size
must include space for the terminator.
Known runtime type classes appear by their TYPE_ names; unknown values retain their decimal codes.
</description>
*)
//!<param name="oldSubstring">Text to replace; empty performs no replacements.</param>
//!<param name="newSubstring">Replacement text; empty deletes each selected match.</param>
//!<param name="replacementCount">Number of completed replacements.</param>
METHOD ReplaceInSource255
VAR_INPUT
	sourceString : ANY_STRING;
	oldSubstring : STRING(255);
	newSubstring : STRING(255);
	maxReplacements : UINT := 0;
	skipReplacements : UINT := 0;
END_VAR
VAR_OUTPUT
	replacementCount : UINT;
END_VAR
VAR	
	
	replaceResult : BOOL; 
END_VAR
VAR
	formattedExceptionMessage : WSTRING(255);
END_VAR
IF sourceString.TypeClass <> __SYSTEM.TYPE_CLASS.TYPE_STRING THEN
	formattedExceptionMessage := Tc2_Utilities.WCONCAT(
		STR1 := "Not supported type ",
		STR2 := SystemTypeClassConvertor.ToWideString(typeClass := sourceString.TypeClass)
	);

	Exceptions.ThrowNotSupported(
		sourceNamespaceName := NamespaceName,
		sourceClassName := ClassName,
		sourcePOUName := __POUNAME(),
		sourcePosition := __POSITION(),
		message := formattedExceptionMessage
	);
END_IF

IF NOT InternalReplaceInSource(
	sourceString := sourceString,
	oldSubstring := ADR(oldSubstring),
	newSubstring := ADR(newSubstring),
	maxReplacements := maxReplacements,
	skipReplacements := skipReplacements,
	replacementCount => replacementCount
) THEN
	Exceptions.ThrowTargetVariableMemoryOverflow(
		sourceNamespaceName := NamespaceName,
		sourceClassName := ClassName,
		sourcePOUName := __POUNAME(),
		sourcePosition := __POSITION(),
		targetVariableName := 'sourceString',
		targetVariableSize := TO_UDINT(sourceString.diSize)
	);
END_IF
END_METHOD

(*!
<summary>Builds a borrowed ANY descriptor for text at an address.</summary>
<description>
Requires a nonzero address to valid terminated text. Records occupied bytes including the terminator, not
buffer capacity; size must fit DINT. Does not copy, allocate or acquire ownership. Keep the source alive while
using the descriptor.
</description>
*)
METHOD StringPointerToAnyType : __System.AnyType
VAR_INPUT
	value : POINTER TO STRING;
END_VAR
StringPointerToAnyType.TypeClass := __SYSTEM.TYPE_CLASS.TYPE_STRING;
StringPointerToAnyType.pValue := value;
StringPointerToAnyType.diSize := TO_DINT(GetActualSize(value^));
END_METHOD

(*!
<summary>Builds a borrowed ANY descriptor for a string reference.</summary>
<description>
Requires a valid reference to terminated text. Records occupied bytes including the terminator, not buffer
capacity; size must fit DINT. Keep the source alive while using the descriptor; no ownership is transferred.
</description>
*)
METHOD StringReferenceToAnyType : __System.AnyType
VAR_INPUT
	value : REFERENCE TO STRING;
END_VAR
StringReferenceToAnyType.TypeClass := __SYSTEM.TYPE_CLASS.TYPE_STRING;
StringReferenceToAnyType.pValue := ADR(value);
StringReferenceToAnyType.diSize := TO_DINT(GetActualSize(value));
END_METHOD

(*!
<summary>Builds a borrowed ANY descriptor for the supplied string.</summary>
<description>
Records occupied bytes including the terminator, not buffer capacity; size must fit DINT. Does not copy or
acquire ownership. Do not retain the descriptor beyond the source lifetime.
</description>
*)
METHOD StringToAnyType : __SYSTEM.AnyType
VAR_IN_OUT CONSTANT
	value : STRING;
END_VAR
StringToAnyType.TypeClass := __SYSTEM.TYPE_CLASS.TYPE_STRING;
StringToAnyType.pValue := ADR(value);
StringToAnyType.diSize := TO_DINT(GetActualSize(value));
END_METHOD

(*!
<summary>Removes repetitions of one character from the selected ends of a string.</summary>
<description>
Modifies the supplied string in place using TrimChars and the requested trim mode. Preserves the remaining
character order and requires writable terminated text.
</description>
*)
METHOD TrimChar
VAR_IN_OUT
	stringToTrim : STRING;
END_VAR
VAR_INPUT
	trimMode : TRIM_MODE := TRIM_MODE.LEFT_AND_RIGHT;
	trimChar : STRING(1) := ' ';
END_VAR
VAR
	trimCharArray : ARRAY [0..0] OF STRING(1);	
END_VAR
trimCharArray[0] := trimChar;

TrimChars(stringToTrim := stringToTrim, trimMode := trimMode, trimChars := trimCharArray);
END_METHOD

(*!
<summary>Removes selected character values from the requested ends of a string in place.</summary>
<description>
The caller supplies a live writable null-terminated string. Left trimming moves the retained suffix, including
its terminator, within the same buffer; no new storage is allocated. The trim-character array may have
negative bounds. Right trimming stops after the first code unit without decrementing an unsigned index below
zero.
</description>
*)
METHOD TrimChars
VAR_IN_OUT
	stringToTrim : STRING;
END_VAR
VAR_INPUT
	trimMode : TRIM_MODE := TRIM_MODE.LEFT_AND_RIGHT;
END_VAR
VAR_IN_OUT CONSTANT
	trimChars : ARRAY [*] OF STRING(1);	
END_VAR
VAR
	stringLength : UDINT;
	stringData : POINTER TO BYTE;
	trimCharData : POINTER TO BYTE;
	
	originalCharIndex : UDINT;
	trimCharIndex : DINT;
	trimCharCount : UDINT;
END_VAR
stringData := ADR(stringToTrim);
stringLength := InternalGetLength(value := stringData);

IF stringLength < 1 THEN
	RETURN;
END_IF

IF trimMode = TRIM_MODE.LEFT_AND_RIGHT OR_ELSE trimMode = TRIM_MODE.LEFT THEN
	trimCharCount := 0;
	
	FOR originalCharIndex := 0 TO stringLength - 1 BY 1 DO
		FOR trimCharIndex := LOWER_BOUND(trimChars, 1) TO UPPER_BOUND(trimChars, 1) DO
			trimCharData := ADR(trimChars[trimCharIndex]);
			
			IF stringData[originalCharIndex] = trimCharData^ THEN
				trimCharCount := trimCharCount + 1;
				EXIT;
			END_IF
		END_FOR
		
		IF trimCharCount <> originalCharIndex + 1 THEN
			EXIT;
		END_IF
	END_FOR

	IF trimCharCount > 0 THEN
		stringLength := stringLength - trimCharCount;
		
		Tc2_System.MEMMOVE(
			destAddr := stringData,
			srcAddr := stringData + (trimCharCount * CharSize),
			n := (stringLength * CharSize) + CharSize
		);		
	END_IF
END_IF

IF stringLength < 1 THEN
	RETURN;
END_IF

IF trimMode = TRIM_MODE.LEFT_AND_RIGHT OR_ELSE trimMode = TRIM_MODE.RIGHT THEN
	trimCharCount := 0;
	
	FOR originalCharIndex := stringLength TO 1 BY -1 DO
		FOR trimCharIndex := LOWER_BOUND(trimChars, 1) TO UPPER_BOUND(trimChars, 1) DO
			trimCharData := ADR(trimChars[trimCharIndex]);
			
			IF stringData[originalCharIndex - 1] = trimCharData^ THEN
				trimCharCount := trimCharCount + 1;
				EXIT;
			END_IF
		END_FOR
		
		IF trimCharCount <> stringLength - originalCharIndex + 1 THEN
			EXIT;
		END_IF
	END_FOR

	IF trimCharCount > 0 THEN
		stringLength := stringLength - trimCharCount;
		
		Tc2_System.MEMSET(destAddr := stringData + (stringLength * CharSize), fillByte := 0, n := CharSize);		
	END_IF	
END_IF
END_METHOD

(*!
<summary>Appends one STRING to a caller-owned buffer and reports success.</summary>
<description>
Requires live, null-terminated source strings and a writable STRING target with valid capacity metadata. Empty
fragments do not stop processing; if all are empty, the target is unchanged and the operation succeeds.
Returns FALSE for a non-STRING target or when appending fails. Processing stops on the first append failure;
earlier modifications are not rolled back. Source storage is borrowed only for this call. Catches exceptions
and returns FALSE; terminal allocation state is preserved for the task boundary. Partial writes are not rolled
back. Valid buffer lifetime and capacity remain caller preconditions.
</description>
*)
METHOD TryAppend : BOOL
VAR_INPUT
	targetString : ANY_STRING;
END_VAR
VAR_IN_OUT CONSTANT
	sourceString : STRING;
END_VAR
__TRY
	TryAppend := InternalAppend(
		targetString := targetString,
		sourceString1 := ADR(sourceString),
		sourceString2 := 0,
		sourceString3 := 0,
		sourceString4 := 0,
		sourceString5 := 0,
		sourceString6 := 0,
		sourceString7 := 0,
		sourceString8 := 0,
		sourceString9 := 0,
		sourceString10 := 0
	);
__CATCH
	TryAppend := FALSE;
__ENDTRY
END_METHOD

(*!
<summary>Appends up to ten STRING fragments in argument order, skipping empty fragments.</summary>
<description>
Requires live, null-terminated source strings and a writable STRING target with valid capacity metadata. Empty
fragments do not stop processing; if all are empty, the target is unchanged and the operation succeeds.
Returns FALSE for a non-STRING target or when appending fails. Processing stops on the first append failure;
earlier modifications are not rolled back. Source storage is borrowed only for this call. Catches exceptions
and returns FALSE; terminal allocation state is preserved for the task boundary. Partial writes are not rolled
back. Valid buffer lifetime and capacity remain caller preconditions.
</description>
*)
METHOD TryAppend255 : BOOL
VAR_INPUT
	targetString : ANY_STRING;
	sourceString1 : STRING(255);
	sourceString2 : STRING(255) := '';
	sourceString3 : STRING(255) := '';
	sourceString4 : STRING(255) := '';
	sourceString5 : STRING(255) := '';
	sourceString6 : STRING(255) := '';
	sourceString7 : STRING(255) := '';
	sourceString8 : STRING(255) := '';
	sourceString9 : STRING(255) := '';
	sourceString10 : STRING(255) := '';
END_VAR
__TRY
	TryAppend255 := InternalAppend(
		targetString := targetString,
		sourceString1 := ADR(sourceString1),
		sourceString2 := ADR(sourceString2),
		sourceString3 := ADR(sourceString3),
		sourceString4 := ADR(sourceString4),
		sourceString5 := ADR(sourceString5),
		sourceString6 := ADR(sourceString6),
		sourceString7 := ADR(sourceString7),
		sourceString8 := ADR(sourceString8),
		sourceString9 := ADR(sourceString9),
		sourceString10 := ADR(sourceString10)
	);
__CATCH
	TryAppend255 := FALSE;
__ENDTRY
END_METHOD

(*!
<summary>Appends text to a STRING buffer, marking truncation when capacity permits.</summary>
<description>
Requires live, terminated input and writable target storage of the matching encoding.
On overflow, capacities of at least three characters use three dots. Capacities of one or two use one dot.
A buffer with room only for its terminator stays empty and succeeds. Missing terminator space or an invalid
target returns FALSE. Exceptions are contained.
</description>
<param name="targetString">Writable STRING buffer to append to.</param>
<param name="sourceString">Text to append; empty leaves the target unchanged.</param>
*)
METHOD TryAppendFit : BOOL
VAR_INPUT
	targetString : ANY_STRING;
END_VAR
VAR_IN_OUT CONSTANT
	sourceString : STRING;
END_VAR
__TRY
	TryAppendFit := InternalAppendFit(targetString := targetString, sourceString := ADR(sourceString));
__CATCH
	TryAppendFit := FALSE;
__ENDTRY
END_METHOD

(*!
<summary>Appends ordered fragments to a STRING buffer, marking truncation when capacity permits.</summary>
<description>
Requires live, terminated input and writable target storage of the matching encoding.
Processes fragments in order. Completed appends remain visible on failure.
On overflow, capacities of at least three characters use three dots. Capacities of one or two use one dot.
A buffer with room only for its terminator stays empty and succeeds. Missing terminator space or an invalid
target returns FALSE. Exceptions are contained.
</description>
<param name="targetString">Writable STRING buffer to append to.</param>
<param name="sourceString1">First text fragment to append.</param>
<param name="sourceString2">Second text fragment to append.</param>
<param name="sourceString3">Third text fragment to append.</param>
<param name="sourceString4">Fourth text fragment to append.</param>
<param name="sourceString5">Fifth text fragment to append.</param>
<param name="sourceString6">Sixth text fragment to append.</param>
<param name="sourceString7">Seventh text fragment to append.</param>
<param name="sourceString8">Eighth text fragment to append.</param>
<param name="sourceString9">Ninth text fragment to append.</param>
<param name="sourceString10">Tenth text fragment to append.</param>
*)
METHOD TryAppendFit255 : BOOL
VAR_INPUT
	targetString : ANY_STRING;
	sourceString1 : STRING(255);
	sourceString2 : STRING(255) := '';
	sourceString3 : STRING(255) := '';
	sourceString4 : STRING(255) := '';
	sourceString5 : STRING(255) := '';
	sourceString6 : STRING(255) := '';
	sourceString7 : STRING(255) := '';
	sourceString8 : STRING(255) := '';
	sourceString9 : STRING(255) := '';
	sourceString10 : STRING(255) := '';
END_VAR
__TRY
	TryAppendFit255 := FALSE;

	IF targetString.TypeClass <> __SYSTEM.TYPE_CLASS.TYPE_STRING THEN
		RETURN;
	END_IF

	IF NOT InternalAppendFit(targetString := targetString, sourceString := ADR(sourceString1)) THEN
		RETURN;
	END_IF

	IF sourceString2 <> '' AND_THEN NOT InternalAppendFit(targetString := targetString, sourceString := ADR(sourceString2)) THEN
		RETURN;
	END_IF

	IF sourceString3 <> '' AND_THEN NOT InternalAppendFit(targetString := targetString, sourceString := ADR(sourceString3)) THEN
		RETURN;
	END_IF

	IF sourceString4 <> '' AND_THEN NOT InternalAppendFit(targetString := targetString, sourceString := ADR(sourceString4)) THEN
		RETURN;
	END_IF

	IF sourceString5 <> '' AND_THEN NOT InternalAppendFit(targetString := targetString, sourceString := ADR(sourceString5)) THEN
		RETURN;
	END_IF

	IF sourceString6 <> '' AND_THEN NOT InternalAppendFit(targetString := targetString, sourceString := ADR(sourceString6)) THEN
		RETURN;
	END_IF

	IF sourceString7 <> '' AND_THEN NOT InternalAppendFit(targetString := targetString, sourceString := ADR(sourceString7)) THEN
		RETURN;
	END_IF

	IF sourceString8 <> '' AND_THEN NOT InternalAppendFit(targetString := targetString, sourceString := ADR(sourceString8)) THEN
		RETURN;
	END_IF

	IF sourceString9 <> '' AND_THEN NOT InternalAppendFit(targetString := targetString, sourceString := ADR(sourceString9)) THEN
		RETURN;
	END_IF

	IF sourceString10 <> '' AND_THEN NOT InternalAppendFit(targetString := targetString, sourceString := ADR(sourceString10)) THEN
		RETURN;
	END_IF

	TryAppendFit255 := TRUE;
__CATCH
	TryAppendFit255 := FALSE;
__ENDTRY
END_METHOD

(*!
<summary>Initializes a splitter when the source has the supported string type.</summary>
<description>
The source must remain alive and unchanged during iteration. The splitter owns its current fragment; borrowed
fragment references expire on MoveNext, Reset or destruction. This method does not allocate the splitter with
__NEW. The initialized result has no fragment allocation until MoveNext; assigning it must not overwrite an
instance with an unreleased fragment. The caller is responsible for the result lifetime and cleanup, including
Reset when abandoning iteration. Do not copy an active splitter by value; use references. Only an instance
explicitly allocated with __NEW may be deleted with __DELETE. Catches exceptions and returns FALSE; terminal
allocation state is preserved for the task boundary. A null source address or missing terminator capacity
returns FALSE before initialization.
Use the output only after TRUE is returned.
</description>
*)
//!<param name="maxCount">
//! Maximum number of returned fragments; zero means unlimited. Empty fragments removed after optional
//! trimming do not count toward the limit. Remaining text is not returned after the limit is reached and is
//! not merged into the last fragment.
//! </param>
//!<param name="separator">
//! Copied separator containing 1 to 80 characters. An invalid reference, empty or longer value returns FALSE
//! before initialization. The 255-character input capacity preserves rejection of all values longer than 80.
//! </param>
METHOD TryCreateSplitter : BOOL
VAR_INPUT
	sourceString : ANY_STRING;
END_VAR
VAR_INPUT
	separator : STRING(255);
	maxCount : UDINT := 0;
	trimEntries : BOOL := FALSE;
	removeEmptyEntries : BOOL := FALSE;
END_VAR
VAR_OUTPUT
	splitter : StringSplittingEnumerator;
END_VAR
__TRY
	IF sourceString.TypeClass <> __SYSTEM.TYPE_CLASS.TYPE_STRING
		OR_ELSE sourceString.pValue = Memory.NULL_ADDRESS
		OR_ELSE sourceString.diSize < TO_DINT(CharSize)
	THEN
		RETURN;
	END_IF

	IF separator = '' OR_ELSE InternalGetLength(value := ADR(separator)) > 80 THEN
		RETURN;
	END_IF

	splitter.Initialize(
		sourceString := sourceString.pValue,
		separator := separator,
		maxCount := maxCount,
		trimEntries := trimEntries,
		removeEmptyEntries := removeEmptyEntries
	);

	TryCreateSplitter := TRUE;
__CATCH
	TryCreateSplitter := FALSE;
__ENDTRY
END_METHOD

(*!
<summary>Joins enumerated values into a caller-owned STRING buffer.</summary>
<description>
Returns FALSE on terminal allocation failure, including when an enumerator catches the original exception.
Borrows and advances the enumerator from its current position. Clears the target before joining; previous
target contents and enumerator position are not restored on failure. Catches exceptions and returns FALSE;
terminal allocation state is preserved for the task boundary. Partial writes are not rolled back. Valid buffer
lifetime and capacity remain caller preconditions.
</description>
*)
METHOD TryJoin : BOOL
VAR_INPUT
	targetString : ANY_STRING;
END_VAR
VAR_INPUT
	separator : STRING;
	sourceEnumerator : IEnumerator;
	startIndex : UDINT := 0;
	count : UDINT := 0;
END_VAR
__TRY
	TryJoin := InternalJoin(
		targetString := targetString,
		separator := ADR(separator),
		sourceEnumerator := sourceEnumerator,
		startIndex := startIndex,
		count := count
	);
__CATCH
	TryJoin := FALSE;
__ENDTRY
END_METHOD

(*!
<summary>Replaces matching substrings in the supplied text buffer.</summary>
<description>
Replaces exact, case-sensitive, non-overlapping occurrences in place. An empty oldSubstring succeeds without
changes and sets replacementCount to zero. An empty newSubstring deletes matched text. Zero maxReplacements
means no replacement limit; skipReplacements skips the first matching occurrences. Returns FALSE for an
incompatible source type or if replacement cannot complete. Replacement is not atomic. If the next replacement
would exceed buffer capacity, it is not performed; completed replacements remain, replacementCount reports
their count, and the valid source remains null-terminated. These guarantees concern capacity failure with
valid input buffers, not invalid memory access. The caller supplies live buffers of the correct encoding;
sourceString must be writable and its size must include space for the terminator. Catches exceptions and
returns FALSE; terminal allocation state is preserved for the task boundary. Partial writes are not rolled
back. Valid buffer lifetime and capacity remain caller preconditions.
</description>
*)
//!<param name="oldSubstring">Text to replace; empty performs no replacements.</param>
//!<param name="newSubstring">Replacement text; empty deletes each selected match.</param>
//!<param name="replacementCount">Number of completed replacements.</param>
METHOD TryReplaceInSource : BOOL
VAR_INPUT
	sourceString : ANY_STRING;
END_VAR
VAR_IN_OUT CONSTANT
	oldSubstring : STRING;
	newSubstring : STRING;
END_VAR
VAR_INPUT
	maxReplacements : UINT := 0;
	skipReplacements : UINT := 0;
END_VAR
VAR_OUTPUT
	replacementCount : UINT;
END_VAR
__TRY
	IF sourceString.TypeClass <> __SYSTEM.TYPE_CLASS.TYPE_STRING THEN
		RETURN;
	END_IF

	TryReplaceInSource := InternalReplaceInSource(
		sourceString := sourceString,
		oldSubstring := ADR(oldSubstring),
		newSubstring := ADR(newSubstring),
		maxReplacements := maxReplacements,
		skipReplacements := skipReplacements,
		replacementCount => replacementCount
	);
__CATCH
	TryReplaceInSource := FALSE;
__ENDTRY
END_METHOD

(*!
<summary>Replaces matching substrings in the supplied text buffer.</summary>
<description>
Replaces exact, case-sensitive, non-overlapping occurrences in place. An empty oldSubstring succeeds without
changes and sets replacementCount to zero. An empty newSubstring deletes matched text. Zero maxReplacements
means no replacement limit; skipReplacements skips the first matching occurrences. Returns FALSE for an
incompatible source type or if replacement cannot complete. Replacement is not atomic. If the next replacement
would exceed buffer capacity, it is not performed; completed replacements remain, replacementCount reports
their count, and the valid source remains null-terminated. These guarantees concern capacity failure with
valid input buffers, not invalid memory access. The caller supplies live buffers of the correct encoding;
sourceString must be writable and its size must include space for the terminator. Catches exceptions and
returns FALSE; terminal allocation state is preserved for the task boundary. Partial writes are not rolled
back. Valid buffer lifetime and capacity remain caller preconditions.
</description>
*)
//!<param name="oldSubstring">Text to replace; empty performs no replacements.</param>
//!<param name="newSubstring">Replacement text; empty deletes each selected match.</param>
//!<param name="replacementCount">Number of completed replacements.</param>
METHOD TryReplaceInSource255 : BOOL
VAR_INPUT
	sourceString : ANY_STRING;
	oldSubstring : STRING(255);
	newSubstring : STRING(255);
	maxReplacements : UINT := 0;
	skipReplacements : UINT := 0;
END_VAR
VAR_OUTPUT
	replacementCount : UINT;
END_VAR
__TRY
	IF sourceString.TypeClass <> __SYSTEM.TYPE_CLASS.TYPE_STRING THEN
		RETURN;
	END_IF

	TryReplaceInSource255 := InternalReplaceInSource(
		sourceString := sourceString,
		oldSubstring := ADR(oldSubstring),
		newSubstring := ADR(newSubstring),
		maxReplacements := maxReplacements,
		skipReplacements := skipReplacements,
		replacementCount => replacementCount
	);
__CATCH
	TryReplaceInSource255 := FALSE;
__ENDTRY
END_METHOD

END_PROGRAM

(* stored: Version 1.1.0.1
   POU Strings: Id {7aa7463a-7b84-4807-b00e-cbaa6fc59270}, SpecialFunc None
   Folder Any: Id {8688dfc3-2927-467c-9f5b-91ce2217a978}
   Folder Append: Id {7e7c80a5-b2b3-4398-aeb3-fcbeeedb95b0}
   Folder Join: Id {23020608-d9f6-4bcd-bc2c-4f5978ed3025}
   Folder Replace: Id {a7f2f348-7292-464d-8aaa-84a00bdb1d6c}
   Folder Service members: Id {6eebbe56-ba8f-4c4e-a22c-3fcf35f9aa27}
   Folder Split: Id {abd107b6-e51f-460b-baa2-99a9483990d2}
   Folder Trim: Id {f20b62c4-34de-4080-969d-424865288d4e}
   Method AnyToString: Id {b226cb15-ac0d-48f7-98b9-48ee0196d1ce}
   Method AnyToString255: Id {6ec6dde0-5575-44dd-bea2-d21349d12524}
   Method AnyToStringFit255: Id {64a20004-3f77-4b1a-908f-282a178d2bc7}
   Method Append: Id {7d3432ad-7058-4ce7-80d2-01c9d35ec6fb}
   Method Append255: Id {b845707e-9f67-4676-b647-f64266f03b85}
   Method AppendFit: Id {64a20001-3f77-4b1a-908f-282a178d2bc7}
   Method AppendFit255: Id {741614c7-882a-4b63-b2d0-ee975117324f}
   Property ClassName: Id {81cda6c2-0106-408d-bf8b-7dd5b920c809}
   Get Get: Id {566edcc0-aa57-4ecd-95d3-18653d40dc60}
   Method Concat255: Id {833ffcb1-3f77-4b1a-908f-282a178d2bc7}
   Method ConcatFit255: Id {64a20003-3f77-4b1a-908f-282a178d2bc7}
   Method Contains: Id {382d5dec-076a-4371-95cd-edb6d9d627f6}
   Method CreateSplitter: Id {74505d39-c9b2-47f5-a8a1-80fe0e3aaae8}
   Method Find: Id {0c61da8f-b806-465e-b4f1-5bdbe54f1092}
   Method GetActualSize: Id {e8e8416f-8e42-44ac-ac9b-ab76e4a16eec}
   Method GetLength: Id {a3dc2c45-cc1a-482d-b619-dbbdf1878690}
   Method InternalAnyToString255: Id {dbd6569e-fd5b-4765-a843-fc6bef815e68}
   Method InternalAppend: Id {96f09b6b-a3b9-4899-b746-36fdcd4d9236}
   Method InternalAppendFit: Id {64a20005-3f77-4b1a-908f-282a178d2bc7}
   Method InternalFind: Id {5b6aff61-016c-4db4-94ed-cfbbb336515e}
   Method InternalGetLength: Id {06d76460-e6eb-42be-8f6b-fb87a2b574a4}
   Method InternalJoin: Id {641619b9-d14d-4e22-94f4-454b0a713080}
   Method InternalReplaceInSource: Id {0ac24766-5e3a-42f7-a2a0-58aa460f844f}
   Method IsFloat: Id {5cca10b4-3ba5-4176-ae1b-a21dca6dbf97}
   Method IsInteger: Id {64017c0a-0904-4813-83bf-5a23b0d4cfee}
   Method IsNullOrWhiteSpace: Id {523b397c-6e9a-4d05-935a-38a2426b04e1}
   Method IsUnsignedInteger: Id {dfaddadb-137b-494a-9d2f-8a9a940574ca}
   Method Join: Id {f9356af7-1c6b-416a-a5c8-0029f23752d3}
   Property NamespaceName: Id {475cd351-78e5-4557-baf1-9d5933c3fa2e}
   Get Get: Id {2b015e66-fd97-4ebe-8516-bd91f7e0b822}
   Method ReplaceInSource: Id {f06898de-32ea-4f51-b053-1b282cb73a8a}
   Method ReplaceInSource255: Id {f41fa253-7b57-4bb9-a052-ea59a6eb6bff}
   Method StringPointerToAnyType: Id {a10ef46f-9469-4b72-b2c7-fdc82174f321}
   Method StringReferenceToAnyType: Id {06b7793c-cb19-41ed-b05e-889daf02c80f}
   Method StringToAnyType: Id {ad63b85b-ddb5-45f3-baef-6d6cd1517473}
   Method TrimChar: Id {62b24a6d-bbc4-486f-b32e-31180d926835}
   Method TrimChars: Id {f8f9620e-29b0-4754-aeb8-6e676ec3c2d0}
   Method TryAppend: Id {bf1d041e-2745-49ca-b076-368f2e842cc8}
   Method TryAppend255: Id {9c82266a-bb32-451c-9763-5118bd999fda}
   Method TryAppendFit: Id {64a20002-3f77-4b1a-908f-282a178d2bc7}
   Method TryAppendFit255: Id {f69b240f-5523-4365-b6d7-898cb6a46d47}
   Method TryCreateSplitter: Id {34df4a0d-a862-4e0c-8436-c7e6b40e8278}
   Method TryJoin: Id {a81f6dab-b206-48bb-a5a8-39b9933d426e}
   Method TryReplaceInSource: Id {6cd9fde4-681b-4169-adb0-283364fff827}
   Method TryReplaceInSource255: Id {9f1f7515-63df-42e0-8ebb-d9a7a98ddbf5} *)
